TYPE E_ErrorFormat :(
	eErrID:=0,
	eErrLevel:=1,
	eErrMeassage:=2,
	eErrModuleDescription:=3
);
END_TYPE

(* stored: Version 1.1.0.1, ProductVersion 3.1.4024.13
   DUT E_ErrorFormat: Id {0b00f3a3-fa79-48b2-81fd-c602943b832e} *)
